TYPE ST_PolarIIChamber_OutsideRingServiceStatus :
STRUCT
	Lift : ST_PolarIIChamber_LiftTopDownServiceStatus;
	Rotate : ST_PolarIIChamber_OutsideRingRotateServiceStatus;
END_STRUCT
END_TYPE

(* stored: Version 1.1.0.1, ProductVersion 3.1.4026.18
   DUT ST_PolarIIChamber_OutsideRingServiceStatus: Id {14000000-0000-0000-0000-000000000069} *)
